Staubli VAL3: Action.dtx

actCmdType actCmd[40]
  [0]
    bool bActFinish
    num nActionID
    num nMoveID
    string sActName
  [1]
    bool bActFinish
    num nActionID
    num nMoveID
    string sActName
  [2]
    bool bActFinish
    num nActionID
    num nMoveID
    string sActName
  [3]
    bool bActFinish
    num nActionID
    num nMoveID
    string sActName
  [4]
    bool bActFinish
    num nActionID
    num nMoveID
    string sActName
  [5]
    bool bActFinish
    num nActionID
    num nMoveID
    string sActName
  [6]
    bool bActFinish
    num nActionID
    num nMoveID
    string sActName
  [7]
    bool bActFinish
    num nActionID
    num nMoveID
    string sActName
  [8]
    bool bActFinish
    num nActionID
    num nMoveID
    string sActName
  [9]
    bool bActFinish
    num nActionID
    num nMoveID
    string sActName
  [10]
    bool bActFinish
    num nActionID
    num nMoveID
    string sActName
  [11]
    bool bActFinish
    num nActionID
    num nMoveID
    string sActName
  [12]
    bool bActFinish
    num nActionID
    num nMoveID
    string sActName
  [13]
    bool bActFinish
    num nActionID
    num nMoveID
    string sActName
  [14]
    bool bActFinish
    num nActionID
    num nMoveID
    string sActName
  [15]
    bool bActFinish
    num nActionID
    num nMoveID
    string sActName
  [16]
    bool bActFinish
    num nActionID
    num nMoveID
    string sActName
  [17]
    bool bActFinish
    num nActionID
    num nMoveID
    string sActName
  [18]
    bool bActFinish
    num nActionID
    num nMoveID
    string sActName
  [19]
    bool bActFinish
    num nActionID
    num nMoveID
    string sActName
  [20]
    bool bActFinish
    num nActionID
    num nMoveID
    string sActName
  [21]
    bool bActFinish
    num nActionID
    num nMoveID
    string sActName
  [22]
    bool bActFinish
    num nActionID
    num nMoveID
    string sActName
  [23]
    bool bActFinish
    num nActionID
    num nMoveID
    string sActName
  [24]
    bool bActFinish
    num nActionID
    num nMoveID
    string sActName
  [25]
    bool bActFinish
    num nActionID
    num nMoveID
    string sActName
  [26]
    bool bActFinish
    num nActionID
    num nMoveID
    string sActName
  [27]
    bool bActFinish
    num nActionID
    num nMoveID
    string sActName
  [28]
    bool bActFinish
    num nActionID
    num nMoveID
    string sActName
  [29]
    bool bActFinish
    num nActionID
    num nMoveID
    string sActName
  [30]
    bool bActFinish
    num nActionID
    num nMoveID
    string sActName
  [31]
    bool bActFinish
    num nActionID
    num nMoveID
    string sActName
  [32]
    bool bActFinish
    num nActionID
    num nMoveID
    string sActName
  [33]
    bool bActFinish
    num nActionID
    num nMoveID
    string sActName
  [34]
    bool bActFinish
    num nActionID
    num nMoveID
    string sActName
  [35]
    bool bActFinish
    num nActionID
    num nMoveID
    string sActName
  [36]
    bool bActFinish
    num nActionID
    num nMoveID
    string sActName
  [37]
    bool bActFinish
    num nActionID
    num nMoveID
    string sActName
  [38]
    bool bActFinish
    num nActionID
    num nMoveID
    string sActName
  [39]
    bool bActFinish
    num nActionID
    num nMoveID
    string sActName
actionIO aActionUsing
  [0]
    num nActIO
    num nActResult
    num nActType
actionIO actPrt[40]
  [0]
    num nActIO
    num nActResult
    num nActType
  [1]
    num nActIO
    num nActResult
    num nActType
  [2]
    num nActIO
    num nActResult
    num nActType
  [3]
    num nActIO
    num nActResult
    num nActType
  [4]
    num nActIO
    num nActResult
    num nActType
  [5]
    num nActIO
    num nActResult
    num nActType
  [6]
    num nActIO
    num nActResult
    num nActType
  [7]
    num nActIO
    num nActResult
    num nActType
  [8]
    num nActIO
    num nActResult
    num nActType
  [9]
    num nActIO
    num nActResult
    num nActType
  [10]
    num nActIO
    num nActResult
    num nActType
  [11]
    num nActIO
    num nActResult
    num nActType
  [12]
    num nActIO
    num nActResult
    num nActType
  [13]
    num nActIO
    num nActResult
    num nActType
  [14]
    num nActIO
    num nActResult
    num nActType
  [15]
    num nActIO
    num nActResult
    num nActType
  [16]
    num nActIO
    num nActResult
    num nActType
  [17]
    num nActIO
    num nActResult
    num nActType
  [18]
    num nActIO
    num nActResult
    num nActType
  [19]
    num nActIO
    num nActResult
    num nActType
  [20]
    num nActIO
    num nActResult
    num nActType
  [21]
    num nActIO
    num nActResult
    num nActType
  [22]
    num nActIO
    num nActResult
    num nActType
  [23]
    num nActIO
    num nActResult
    num nActType
  [24]
    num nActIO
    num nActResult
    num nActType
  [25]
    num nActIO
    num nActResult
    num nActType
  [26]
    num nActIO
    num nActResult
    num nActType
  [27]
    num nActIO
    num nActResult
    num nActType
  [28]
    num nActIO
    num nActResult
    num nActType
  [29]
    num nActIO
    num nActResult
    num nActType
  [30]
    num nActIO
    num nActResult
    num nActType
  [31]
    num nActIO
    num nActResult
    num nActType
  [32]
    num nActIO
    num nActResult
    num nActType
  [33]
    num nActIO
    num nActResult
    num nActType
  [34]
    num nActIO
    num nActResult
    num nActType
  [35]
    num nActIO
    num nActResult
    num nActType
  [36]
    num nActIO
    num nActResult
    num nActType
  [37]
    num nActIO
    num nActResult
    num nActType
  [38]
    num nActIO
    num nActResult
    num nActType
  [39]
    num nActIO
    num nActResult
    num nActType
bool bPushToStack
public num _nActStackIndex
num _nNextId
public num _nPuleStartClk[128]
public num nMoveIDRef
num nMoveIdMax = 100
num nSyncMoveID
